Fanuc KAREL source: KT00147.KL

PROGRAM KT00147
%NOLOCKGROUP
VAR
  Y1: ARRAY[2] OF BYTE
  R2: REAL
  OUT: INTEGER
BEGIN
  Y1[1] = 2
    R2 = 3.0
  OUT = Y1[1] DIV R2
END KT00147
